(* LS Electric XG5000 project: TCPUHN *)
(* PLC LSPLC *)

PROGRAM NativeST (* task: 스캔 프로그램 *)
VAR RETAIN
    Count : INT := 7;
END_VAR
VAR
    Delay : TON;
    Message : STRING := 'Ready';
    Samples : ARRAY[0..3] OF INT;
END_VAR
Count := Count + 1;
Samples[0] := Count;
Delay(IN := TRUE, PT := T#1s);
%MX0 := Delay.Q;
Message := 'Running';
END_PROGRAM

PROGRAM NativeIL (* task: 스캔 프로그램 *)
VAR
    Count : INT;
END_VAR
LD 2
ST Count
END_PROGRAM

PROGRAM CreatedST (* task: 스캔 프로그램 *)
VAR RETAIN
    Count : INT := 7;
END_VAR
VAR
    Delay : TON;
    Message : STRING := 'Ready';
    Samples : ARRAY[0..3] OF INT;
END_VAR
Count := Count + 1;
Samples[0] := Count;
Delay(IN := TRUE, PT := T#1s);
%MX0 := Delay.Q;
Message := 'Running';
END_PROGRAM

PROGRAM CreatedIL (* task: 스캔 프로그램 *)
VAR
    Count : INT;
END_VAR
LD 2
ST Count
END_PROGRAM